Fanuc KAREL source: KO00120.KL

PROGRAM KO00120
%NOLOCKGROUP
VAR
  A: ARRAY[2] OF BYTE
  B: ARRAY[2] OF SHORT
  OUT: REAL
BEGIN
  A[1] = 1
  B[1] = 2
  OUT = ATAN2(A[1], B[1])
END KO00120
